FUNCTION_BLOCK Station1Coord (* Basic Function Block Type *)
  (* Standard: 61499-2 *)
  (* Version 0.0, 11/25/2026, Schneider Electric, Station 1 (Distribution + Testing) to Conveyor Stop 1 sequential coordinator *)
  PACKAGE Main;
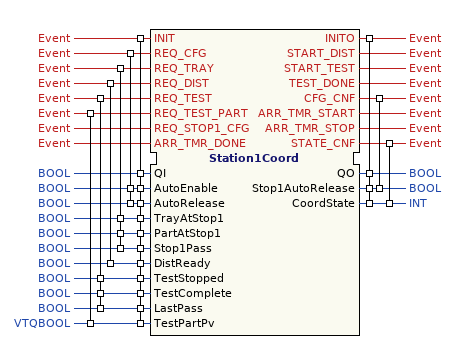
  EVENT_INPUT
    INIT WITH QI, AutoEnable, AutoRelease, TrayAtStop1, PartAtStop1, Stop1Pass, DistReady, TestStopped, TestComplete, LastPass, TestPartPv; (* Initialization Request *)
    REQ_CFG WITH AutoEnable, AutoRelease; (* AutoEnable or AutoRelease toggle update *)
    REQ_TRAY WITH TrayAtStop1, PartAtStop1, Stop1Pass; (* Stop 1 tray and workpiece sensor update *)
    REQ_DIST WITH DistReady; (* Distribution ready state update *)
    REQ_TEST WITH TestStopped, TestComplete, LastPass; (* Testing cycle state and pass/reject result update *)
    REQ_TEST_PART WITH TestPartPv; (* Testing PartAvailable sensor update *)
    REQ_STOP1_CFG; (* Re-emit Stop1AutoRelease config on Conveyor startup *)
    ARR_TMR_DONE; (* Tray arrival settle timer elapsed *)
  END_EVENT
  EVENT_OUTPUT
    INITO WITH QO, Stop1AutoRelease, CoordState; (* Initialization Confirm *)
    START_DIST; (* Start Distribution automatic cycle *)
    START_TEST; (* Start Testing automatic cycle after Distribution has returned home and parked *)
    TEST_DONE; (* Primary Testing pass-complete notification to Conveyor Stop 1 *)
    CFG_CNF WITH Stop1AutoRelease; (* Stop 1 auto-release configuration update *)
    ARR_TMR_START; (* Start tray arrival settle debounce timer *)
    ARR_TMR_STOP; (* Cancel tray arrival settle debounce timer *)
    STATE_CNF WITH CoordState; (* Coordinator state update *)
  END_EVENT
  VAR_INPUT
    QI : BOOL := TRUE; (* Input event qualifier *)
    AutoEnable : BOOL := FALSE; (* Automatic Station 1 mode enable *)
    AutoRelease : BOOL := TRUE; (* Auto-release Stop 1 when filled/passing *)
    TrayAtStop1 : BOOL := FALSE; (* Tray present at Stop 1 (M1.DI02) *)
    PartAtStop1 : BOOL := FALSE; (* Workpiece in Station 1 tray pocket (M1.DI05) *)
    Stop1Pass : BOOL := FALSE; (* Stopper 1 pass-through or releasing state (TRUE=Down, FALSE=Up/Blocking) *)
    DistReady : BOOL := FALSE; (* Distribution CycleSeq Stopped or Completed *)
    TestStopped : BOOL := TRUE; (* Testing CycleSeq Stopped state *)
    TestComplete : BOOL := FALSE; (* Testing CycleSeq Completed state *)
    LastPass : BOOL := FALSE; (* TRUE if last Testing cycle took the pass branch *)
    TestPartPv : VTQBOOL; (* Testing PartAvailable sensor process value *)
  END_VAR
  VAR_OUTPUT
    QO : BOOL; (* Output event qualifier *)
    Stop1AutoRelease : BOOL := FALSE; (* Effective Stop 1 auto-release enable (AutoEnable AND AutoRelease) *)
    CoordState : INT := 0; (* 0=Idle,1=SettleWait,2=RunningDist,3=RunningTest,4=WaitTrayLeave *)
  END_VAR
  VAR
    state : INT := 0; (* Internal state machine value *)
    traySettled : BOOL := FALSE; (* Tray debounce settled at Stop 1 *)
    seenDistRun : BOOL := FALSE; (* Observed Distribution CycleSeq Running since START_DIST *)
    seenTestRun : BOOL := FALSE; (* Observed Testing CycleSeq Running since START_TEST *)
    skipIdle : BOOL := FALSE; (* Prevent same-scan restart after manual Stop *)
    wantStartDist : BOOL := FALSE; (* Pending START_DIST event flag *)
    wantStartTest : BOOL := FALSE; (* Pending START_TEST event flag *)
    wantTestDone : BOOL := FALSE; (* Pending TEST_DONE event flag *)
    wantCfgCnf : BOOL := FALSE; (* Pending CFG_CNF event flag *)
    wantArrStart : BOOL := FALSE; (* Pending ARR_TMR_START event flag *)
    wantArrStop : BOOL := FALSE; (* Pending ARR_TMR_STOP event flag *)
  END_VAR
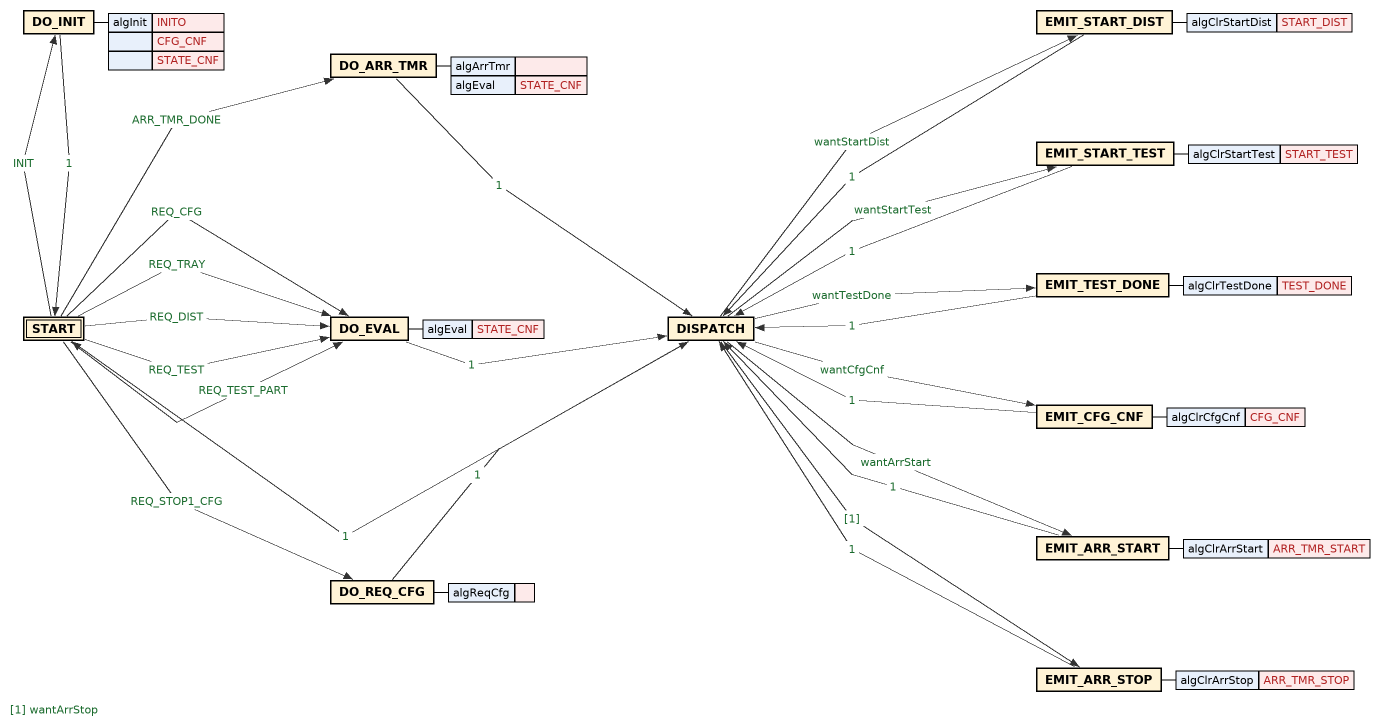
  EC_STATES
    START; (* Initial State *)
    DO_INIT : algInit -> INITO, -> CFG_CNF, -> STATE_CNF;
    DO_EVAL : algEval -> STATE_CNF;
    DO_ARR_TMR : algArrTmr, algEval -> STATE_CNF;
    DO_REQ_CFG : algReqCfg;
    DISPATCH;
    EMIT_START_DIST : algClrStartDist -> START_DIST;
    EMIT_START_TEST : algClrStartTest -> START_TEST;
    EMIT_TEST_DONE : algClrTestDone -> TEST_DONE;
    EMIT_CFG_CNF : algClrCfgCnf -> CFG_CNF;
    EMIT_ARR_START : algClrArrStart -> ARR_TMR_START;
    EMIT_ARR_STOP : algClrArrStop -> ARR_TMR_STOP;
  END_STATES
  EC_TRANSITIONS
    START TO DO_INIT := INIT;
    DO_INIT TO START := 1;
    START TO DO_EVAL := REQ_CFG;
    START TO DO_EVAL := REQ_TRAY;
    START TO DO_EVAL := REQ_DIST;
    START TO DO_EVAL := REQ_TEST;
    START TO DO_EVAL := REQ_TEST_PART;
    START TO DO_ARR_TMR := ARR_TMR_DONE;
    START TO DO_REQ_CFG := REQ_STOP1_CFG;
    DO_EVAL TO DISPATCH := 1;
    DO_ARR_TMR TO DISPATCH := 1;
    DO_REQ_CFG TO DISPATCH := 1;
    DISPATCH TO EMIT_START_DIST := wantStartDist;
    EMIT_START_DIST TO DISPATCH := 1;
    DISPATCH TO EMIT_START_TEST := wantStartTest;
    EMIT_START_TEST TO DISPATCH := 1;
    DISPATCH TO EMIT_TEST_DONE := wantTestDone;
    EMIT_TEST_DONE TO DISPATCH := 1;
    DISPATCH TO EMIT_CFG_CNF := wantCfgCnf;
    EMIT_CFG_CNF TO DISPATCH := 1;
    DISPATCH TO EMIT_ARR_START := wantArrStart;
    EMIT_ARR_START TO DISPATCH := 1;
    DISPATCH TO EMIT_ARR_STOP := wantArrStop;
    EMIT_ARR_STOP TO DISPATCH := 1;
    DISPATCH TO START := 1;
  END_TRANSITIONS
  ALGORITHM algInit IN ST: (* Initialize coordinator state and outputs *)
QO := QI;
state := 0;
traySettled := FALSE;
seenDistRun := FALSE;
seenTestRun := FALSE;
skipIdle := FALSE;
Stop1AutoRelease := AutoEnable AND AutoRelease;
CoordState := 0;
wantStartDist := FALSE;
wantStartTest := FALSE;
wantTestDone := FALSE;
wantCfgCnf := FALSE;
wantArrStart := FALSE;
wantArrStop := FALSE;
  END_ALGORITHM
  ALGORITHM algArrTmr IN ST: (* Mark tray arrival settled when debounce timer expires *)
IF state = 1 THEN
	traySettled := TrayAtStop1 AND (NOT Stop1Pass);
	state := 0;
END_IF;
  END_ALGORITHM
  ALGORITHM algReqCfg IN ST: (* Re-emit Stop1AutoRelease config on Conveyor startup *)
Stop1AutoRelease := AutoEnable AND AutoRelease;
wantCfgCnf := TRUE;
  END_ALGORITHM
  ALGORITHM algEval IN ST: (* Evaluate sequential Station 1 coordination state machine *)
skipIdle := FALSE;

IF Stop1AutoRelease <> (AutoEnable AND AutoRelease) THEN
	Stop1AutoRelease := AutoEnable AND AutoRelease;
	wantCfgCnf := TRUE;
END_IF;

IF NOT AutoEnable THEN
	IF state = 1 THEN
		wantArrStop := TRUE;
	END_IF;
	seenDistRun := FALSE;
	seenTestRun := FALSE;
	state := 0;
ELSE
	IF NOT TrayAtStop1 THEN
		traySettled := FALSE;
		IF state = 1 THEN
			wantArrStop := TRUE;
			state := 0;
		ELSIF state = 4 THEN
			state := 0;
		END_IF;
	ELSIF Stop1Pass THEN
		(* Stopper 1 is down (releasing or Pass mode): cancel settle and never start on passing tray *)
		IF state = 1 THEN
			wantArrStop := TRUE;
			traySettled := FALSE;
			state := 0;
		ELSIF state = 0 THEN
			traySettled := FALSE;
		END_IF;
	END_IF;

	IF state = 2 THEN
		(* RunningDist: wait for Distribution AutoCycle to deliver, return home & park *)
		IF NOT DistReady THEN
			seenDistRun := TRUE;
		ELSIF seenDistRun AND DistReady THEN
			seenDistRun := FALSE;
			IF TestPartPv.value AND (TestStopped OR TestComplete) THEN
				seenTestRun := FALSE;
				wantStartTest := TRUE;
				state := 3;
			ELSE
				state := 0;
				skipIdle := TRUE;
			END_IF;
		END_IF;
	ELSIF state = 3 THEN
		(* RunningTest: wait for TestingCycle pass or reject *)
		IF (NOT TestStopped) AND (NOT TestComplete) THEN
			seenTestRun := TRUE;
		ELSIF seenTestRun AND TestComplete THEN
			seenTestRun := FALSE;
			IF LastPass THEN
				wantTestDone := TRUE;
				IF TrayAtStop1 THEN
					state := 4;
				ELSE
					state := 0;
				END_IF;
			ELSE
				(* Rejected workpiece -> retry on same settled empty tray *)
				state := 0;
			END_IF;
		ELSIF seenTestRun AND TestStopped THEN
			seenTestRun := FALSE;
			state := 0;
			skipIdle := TRUE;
		END_IF;
	END_IF;

	IF (state = 0) AND (NOT skipIdle) AND TrayAtStop1 AND (NOT Stop1Pass) THEN
		IF NOT traySettled THEN
			wantArrStart := TRUE;
			state := 1;
		ELSIF PartAtStop1 THEN
			(* Pre-filled tray: latch WaitTrayLeave so DI05 dropping while leaving never triggers Station 1 *)
			state := 4;
		ELSIF DistReady AND (TestStopped OR TestComplete) THEN
			IF TestPartPv.value THEN
				(* Leftover workpiece already on Testing lift -> test it first *)
				seenTestRun := FALSE;
				wantStartTest := TRUE;
				state := 3;
			ELSE
				seenDistRun := FALSE;
				wantStartDist := TRUE;
				state := 2;
			END_IF;
		END_IF;
	END_IF;
END_IF;

CoordState := state;
  END_ALGORITHM
  ALGORITHM algClrStartDist IN ST: (* Clear START_DIST emit flag *)
wantStartDist := FALSE;
  END_ALGORITHM
  ALGORITHM algClrStartTest IN ST: (* Clear START_TEST emit flag *)
wantStartTest := FALSE;
  END_ALGORITHM
  ALGORITHM algClrTestDone IN ST: (* Clear TEST_DONE emit flag *)
wantTestDone := FALSE;
  END_ALGORITHM
  ALGORITHM algClrCfgCnf IN ST: (* Clear CFG_CNF emit flag *)
wantCfgCnf := FALSE;
  END_ALGORITHM
  ALGORITHM algClrArrStart IN ST: (* Clear ARR_TMR_START emit flag *)
wantArrStart := FALSE;
  END_ALGORITHM
  ALGORITHM algClrArrStop IN ST: (* Clear ARR_TMR_STOP emit flag *)
wantArrStop := FALSE;
  END_ALGORITHM
END_FUNCTION_BLOCK
